INTERFACE I_Gyro

METHOD StartBiasCalibration
END_METHOD

PROPERTY YawRateInRadPerS : LREAL
GET
END_GET
END_PROPERTY

PROPERTY AngularRateInRadPerS : Vector3
GET
END_GET
END_PROPERTY

PROPERTY TimestampInNs : ULINT
GET
END_GET
END_PROPERTY

PROPERTY IsValid : BOOL
GET
END_GET
END_PROPERTY

END_INTERFACE

(* stored: Version 1.1.0.1, ProductVersion 3.1.4026.12
   Itf I_Gyro: Id {d341f671-4619-5705-a9b9-dfbaa4ce28e6}
   Method StartBiasCalibration: Id {a20645ba-519b-593b-91ad-e62ec84239fa}
   Property YawRateInRadPerS: Id {e7a7bfb5-fc38-5d8c-b307-bc14ecd30523}
   Get Get: Id {ccd2e0be-13a5-5aac-9f6f-90cc330f9791}
   Property AngularRateInRadPerS: Id {100af6f7-68bc-5735-9b00-36eac534f159}
   Get Get: Id {33af71ea-99f6-5bf6-9077-9c04c36b553a}
   Property TimestampInNs: Id {c32d565e-3304-5161-a069-c926e6250203}
   Get Get: Id {ad33d0e5-d959-595e-b27f-c39567225e94}
   Property IsValid: Id {e977ceac-fb9d-5a04-80ff-c5d284d9b4e8}
   Get Get: Id {69562f4f-4448-557d-9107-bf7754cdf328} *)
